(* Two Tank Control, One Heating, One Cooling *)

PROGRAM main
  VAR
    Start AT %IX0.0 : BOOL; (* Simple Push Button Input *)
    Stop AT %IX0.1 : BOOL; (* Simple Push Button Input *)
    LevelSensor1 AT %IX0.2 : BOOL;
    LevelSensor2 AT %IX0.3 : BOOL; (* Tank 1 Sensor *)
    LevelSensor3 AT %IX0.4 : BOOL; (* Tank 2 Sensor *)
    LevelSensor4 AT %IX0.5 : BOOL; (* Tank 2 Sensor *)
    CycleOn AT %QX0.0 : BOOL; (* Internal Variable / Output Lamp *)
    InletValve AT %QX0.1 : BOOL; (* Main Inlet Valve Shared by 2 Tanks *)
    Valve2 AT %QX0.2 : BOOL; (* Auxiliary Valve *)
    Valve3 AT %QX0.7 : BOOL; (* Auxiliary Valve *)
    OutletValve1 AT %QX0.3 : BOOL; (* Tank 1 Outlet Valve *)
    OutletValve2 AT %QX0.4 : BOOL; (* Tank 2 Outlet Valve *)
    Heater AT %QX0.5 : BOOL; (* Tank 1 Heater *)
    Cooler AT %QX0.6 : BOOL; (* Tank 2 Cooling Water Flow *)
    TempSensor1 AT %IW1 : INT; (* Tank 1 Analog Temperature Sensor *)
    TempSensor2 AT %IW2 : INT; (* Tank 2 Analog Temperature Sensor *)
  END_VAR

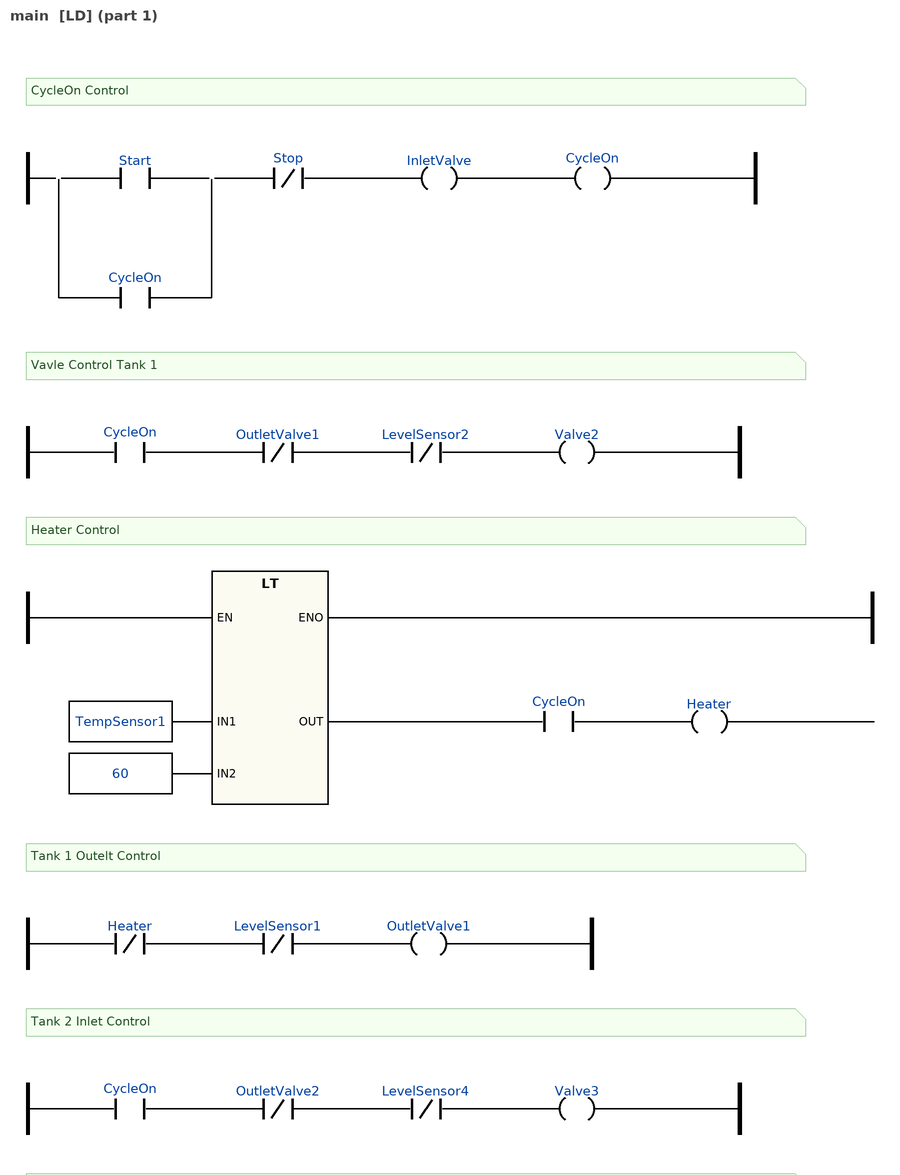
(* LD diagram, written out as Structured Text *)
(* CycleOn Control *)
InletValve := (Start OR CycleOn) AND NOT Stop;
CycleOn := (Start OR CycleOn) AND NOT Stop;
(* Vavle Control Tank 1 *)
Valve2 := CycleOn AND NOT OutletValve1 AND NOT LevelSensor2;
(* Heater Control *)
Heater := TempSensor1 < 60 AND CycleOn;
(* Tank 1 Outelt Control *)
OutletValve1 := NOT Heater AND NOT LevelSensor1;
(* Tank 2 Inlet Control *)
Valve3 := CycleOn AND NOT OutletValve2 AND NOT LevelSensor4;
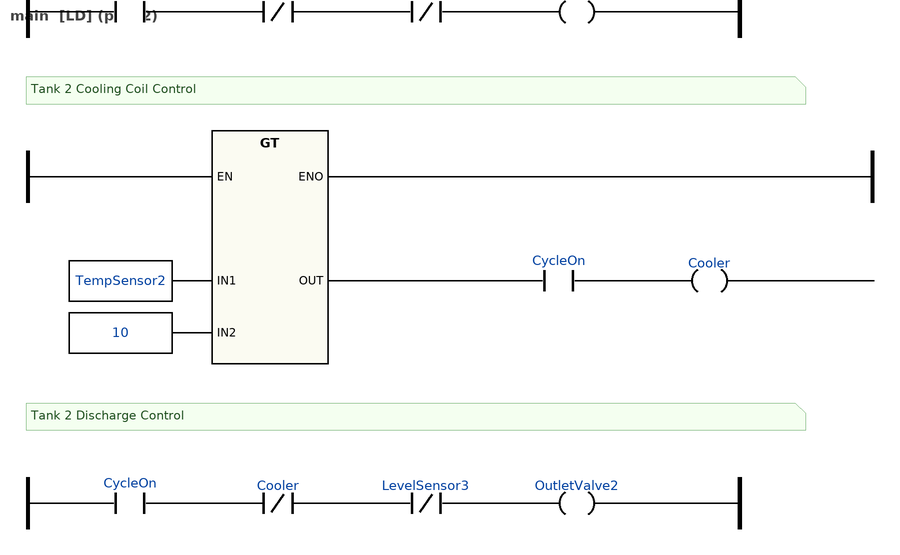
(* Tank 2 Cooling Coil Control *)
Cooler := TempSensor2 > 10 AND CycleOn;
(* Tank 2 Discharge Control *)
OutletValve2 := CycleOn AND NOT Cooler AND NOT LevelSensor3;
END_PROGRAM
